// Model of the TwinSAFE FB TON (switch-on delay).
// The Safety Editor refuses a TON with TonIn1 unconnected: the model then reports Error with diagnostic
// bit 15 instead of running (see T_SafeFunctionBlockBase).
{attribute 'reflection'}
FUNCTION_BLOCK T_SafeTon EXTENDS T_SafeFunctionBlockBase
VAR_INPUT
    TonIn1 : BOOL;
    Parameters : ST_SafeTimerParameters;
END_VAR
VAR_OUTPUT
    TonOut : BOOL;
END_VAR
VAR
    {attribute 'is_connected' := 'TonIn1'}
    _tonIn1Connected : BOOL;
    _state : E_SafeTonState := E_SafeTonState.Stop;
    _timer : TON;
END_VAR

SUPER^();

// TonIn1 must be connected (Safety Editor: "Inport TonIn1 of TON must be connected").
METHOD PROTECTED ConfigurationOk : BOOL
IF NOT _tonIn1Connected THEN
    _configurationFault := 'T_SafeTon: Inport TonIn1 of TON must be connected';
    RETURN;
END_IF

ConfigurationOk := TRUE;
END_METHOD

METHOD PROTECTED Process
VAR
    inputActive : BOOL;
END_VAR
inputActive := _fbRun AND F_SafeInputValue(_tonIn1Connected, Parameters.MakeContact, TonIn1);
_timer(IN := inputActive, PT := Parameters.DelayTime);

IF NOT _fbRun THEN
    _state := E_SafeTonState.Stop;
ELSIF NOT inputActive THEN
    _state := E_SafeTonState.Safe;
ELSIF _timer.Q THEN
    _state := E_SafeTonState.Run;
ELSE
    _state := E_SafeTonState.DelayIn;
END_IF

TonOut := (_state = E_SafeTonState.Run);
Error  := FALSE;
Diag   := 0;
State  := TO_BYTE(_state);
END_METHOD

END_FUNCTION_BLOCK

(* stored: Version 1.1.0.1
   POU T_SafeTon: Id {1b95320b-0d3a-5923-8ff0-0651093a6525}, SpecialFunc None
   Method ConfigurationOk: Id {1e78c1dc-bac7-480d-a034-28eb147ef6d8}
   Method Process: Id {e4417956-7233-5c5f-80ff-76deef0eb2c0} *)
